(****************************************************************************************************<br>
© Syntegon Group.<br>
All rights reserved, also regarding any disposal, exploitation, reproduction, editing, distribution,<br>
as well as in the event of applications for industrial property rights.<br>
*****************************************************************************************************<br>
DESCRIPTION:<br>
Sets pose, track, strokes, gripper offsets and mover size. TRUE if anything changed.<br>
****************************************************************************************************)
METHOD m_Configure : BOOL
VAR_INPUT
	vi_Pose								: ST_VisuPose;	// MCS, track start on top of the movers with Z = 0
	vi_un_ModuleCount					: UINT;	// [-] track modules in a row
	vi_lr_ModuleLength					: LREAL;	// [mm]
	vi_lr_XMin							: LREAL;	// [mm]
	vi_lr_XMax							: LREAL;	// [mm]
	vi_lr_ZMin							: LREAL;	// [mm]
	vi_lr_ZMax							: LREAL;	// [mm]
	vi_lr_ToolOffsetX					: LREAL;	// [mm] gripper flange ahead of the X axis zero
	vi_lr_ToolOffsetZ					: LREAL;	// [mm] gripper flange relative to the mover top (below: negative)
	vi_lr_MoverLength					: LREAL;	// [mm] along the track
	vi_lr_MoverWidth					: LREAL;	// [mm]
END_VAR
VAR
	TempNew								: ST_VisuXtsGantryConfig;
END_VAR
TempNew := vo_Visu.stConfig;
TempNew.stPose := vi_Pose;
TempNew.nModuleCount := vi_un_ModuleCount;
TempNew.fModuleLength := vi_lr_ModuleLength;
TempNew.fXMin := vi_lr_XMin;
TempNew.fXMax := vi_lr_XMax;
TempNew.fZMin := vi_lr_ZMin;
TempNew.fZMax := vi_lr_ZMax;
TempNew.fToolOffsetX := vi_lr_ToolOffsetX;
TempNew.fToolOffsetZ := vi_lr_ToolOffsetZ;
TempNew.fMoverLength := vi_lr_MoverLength;
TempNew.fMoverWidth := vi_lr_MoverWidth;
m_Configure := m_ApplyConfig(TempNew);
END_METHOD

(****************************************************************************************************<br>
© Syntegon Group.<br>
All rights reserved, also regarding any disposal, exploitation, reproduction, editing, distribution,<br>
as well as in the event of applications for industrial property rights.<br>
*****************************************************************************************************<br>
DESCRIPTION:<br>
Sets or clears the fault of the whole gantry: drawn red with the message while active. Faults of single<br>
movers go through m_SetMover. The fault stays until it is cleared with m_SetFault(vi_b_Active := FALSE,<br>
vi_str_Message := ''). TRUE.<br>
****************************************************************************************************)
METHOD m_SetFault : BOOL
VAR_INPUT
	vi_b_Active							: BOOL;	// TRUE: fault active
	vi_str_Message						: STRING(80);	// shown to the operator; empty shows 'Fault'
END_VAR
vo_Visu.stState.stFault.bActive := vi_b_Active;
vo_Visu.stState.stFault.sMessage := vi_str_Message;
m_SetFault := TRUE;
END_METHOD

(****************************************************************************************************<br>
© Syntegon Group.<br>
All rights reserved, also regarding any disposal, exploitation, reproduction, editing, distribution,<br>
as well as in the event of applications for industrial property rights.<br>
*****************************************************************************************************<br>
DESCRIPTION:<br>
Defines finger vi_un_Finger (1-based) of every mover's gripper: a cylinder hanging from the finger's pose along<br>
its local -Z. The finger count grows to vi_un_Finger.<br>
*****************************************************************************************************<br>
OUTPUT VALUES:<br>
FALSE outside 1..VISU_GlobalConst_Param.VISU_un_MAX_FINGERS.<br>
****************************************************************************************************)
METHOD m_SetFinger : BOOL
VAR_INPUT
	vi_un_Finger						: UINT;	// [-] 1-based, as a product's nFingerId
	vi_lr_Diameter						: LREAL;	// [mm]
	vi_lr_Height						: LREAL;	// [mm] along the finger's local -Z
END_VAR
VAR
	TempNew								: ST_VisuXtsGantryConfig;
END_VAR
m_SetFinger := FALSE;
IF vi_un_Finger = 0 OR vi_un_Finger > VISU_GlobalConst_Param.VISU_un_MAX_FINGERS THEN
	RETURN;
END_IF
TempNew := vo_Visu.stConfig;
TempNew.aFingers[vi_un_Finger - 1].fDiameter := vi_lr_Diameter;
TempNew.aFingers[vi_un_Finger - 1].fHeight := vi_lr_Height;
TempNew.nFingerCount := MAX(TempNew.nFingerCount, vi_un_Finger);
m_ApplyConfig(TempNew);
m_SetFinger := TRUE;
END_METHOD

(****************************************************************************************************<br>
© Syntegon Group.<br>
All rights reserved, also regarding any disposal, exploitation, reproduction, editing, distribution,<br>
as well as in the event of applications for industrial property rights.<br>
*****************************************************************************************************<br>
DESCRIPTION:<br>
Reports one mover (actual values) at entry vi_un_Index and marks it valid. Call once per cycle per mover.<br>
*****************************************************************************************************<br>
OUTPUT VALUES:<br>
FALSE if vi_un_Index is outside the mover count set by m_SetMoverCount.<br>
****************************************************************************************************)
METHOD m_SetMover : BOOL
VAR_INPUT
	vi_un_Index							: UINT;	// [-] 0..m_SetMoverCount - 1
	vi_udn_Id							: UDINT;	// [-] unique within the gantry, > 0
	vi_lr_Position						: LREAL;	// [mm] along the track
	vi_lr_X								: LREAL;	// [mm] X axis
	vi_b_GripperActive					: BOOL;	// used only when no fingers are configured
	(* Finger poses absolute in the MCS and grip states, index 0 = finger 1; entries beyond the finger count are ignored. *)
	vi_FingerStates						: ARRAY[0..VISU_GlobalConst_Param.VISU_un_MAX_FINGERS - 1] OF ST_VisuFingerState;
	vi_b_Fault							: BOOL := FALSE;	// TRUE: this mover is in a fault
	vi_str_FaultMessage					: STRING(80) := '';	// shown to the operator; empty shows 'Fault'
END_VAR
m_SetMover := vi_un_Index < vo_Visu.stState.nMoverCount;
IF m_SetMover THEN
	vo_Visu.stState.aMovers[vi_un_Index].nId := vi_udn_Id;
	vo_Visu.stState.aMovers[vi_un_Index].bValid := TRUE;
	vo_Visu.stState.aMovers[vi_un_Index].fPosition := vi_lr_Position;
	vo_Visu.stState.aMovers[vi_un_Index].fX := vi_lr_X;
	vo_Visu.stState.aMovers[vi_un_Index].bGripperActive := vi_b_GripperActive;
	vo_Visu.stState.aMovers[vi_un_Index].aFingerStates := vi_FingerStates;
	vo_Visu.stState.aMovers[vi_un_Index].stFault.bActive := vi_b_Fault;
	vo_Visu.stState.aMovers[vi_un_Index].stFault.sMessage := vi_str_FaultMessage;
	vo_Visu.stState.nTimestamp := m_DcTime();
END_IF
END_METHOD

(****************************************************************************************************<br>
© Syntegon Group.<br>
All rights reserved, also regarding any disposal, exploitation, reproduction, editing, distribution,<br>
as well as in the event of applications for industrial property rights.<br>
*****************************************************************************************************<br>
DESCRIPTION:<br>
Sets how many mover entries are evaluated (limited to VISU_GlobalConst_Param.VISU_un_MAX_MOVERS); entries<br>
beyond are invalidated. TRUE if vi_un_Count fitted.<br>
****************************************************************************************************)
METHOD m_SetMoverCount : BOOL
VAR_INPUT
	vi_un_Count							: UINT;	// [-] movers
END_VAR
VAR
	un_TempIndex						: UINT;
END_VAR
m_SetMoverCount := vi_un_Count <= VISU_GlobalConst_Param.VISU_un_MAX_MOVERS;
vo_Visu.stState.nMoverCount := MIN(vi_un_Count, VISU_GlobalConst_Param.VISU_un_MAX_MOVERS);
FOR un_TempIndex := vo_Visu.stState.nMoverCount TO VISU_GlobalConst_Param.VISU_un_MAX_MOVERS - 1 DO
	vo_Visu.stState.aMovers[un_TempIndex].bValid := FALSE;
END_FOR
END_METHOD

(****************************************************************************************************<br>
© Syntegon Group.<br>
All rights reserved, also regarding any disposal, exploitation, reproduction, editing, distribution,<br>
as well as in the event of applications for industrial property rights.<br>
*****************************************************************************************************<br>
DESCRIPTION:<br>
Moves the gantry's shown coordinate system (origin triad, local measuring coordinates) away from the track<br>
start (stPose), in the gantry's local frame. Geometry and mover positions stay relative to stPose.<br>
TRUE if anything changed.<br>
****************************************************************************************************)
METHOD m_SetOriginShift : BOOL
VAR_INPUT
	vi_lr_X								: LREAL;	// [mm] along the gantry's local X
	vi_lr_Y								: LREAL := 0;	// [mm] along the track (local Y)
	vi_lr_Z								: LREAL := 0;	// [mm] along the gantry's local Z
END_VAR
VAR
	TempNew								: ST_VisuXtsGantryConfig;
END_VAR
TempNew := vo_Visu.stConfig;
TempNew.stOriginShift.fX := vi_lr_X;
TempNew.stOriginShift.fY := vi_lr_Y;
TempNew.stOriginShift.fZ := vi_lr_Z;
m_SetOriginShift := m_ApplyConfig(TempNew);
END_METHOD

(****************************************************************************************************<br>
© Syntegon Group.<br>
All rights reserved, also regarding any disposal, exploitation, reproduction, editing, distribution,<br>
as well as in the event of applications for industrial property rights.<br>
*****************************************************************************************************<br>
DESCRIPTION:<br>
Adds a pick or place zone, or updates the one for the same conveyor and kind.<br>
*****************************************************************************************************<br>
OUTPUT VALUES:<br>
FALSE for vi_udn_ConveyorId = 0 or a full list.<br>
****************************************************************************************************)
METHOD m_SetZone : BOOL
VAR_INPUT
	vi_udn_ConveyorId					: UDINT;	// [-] manifest id of the conveyor
	vi_e_Kind							: E_VisuZoneKind;
	vi_lr_Start							: LREAL;	// [mm] along the conveyor from its origin (belt coordinates, not MCS)
	vi_lr_End							: LREAL;	// [mm] along the conveyor from its origin
	vi_lr_AllocationOffset				: LREAL := 0;	// [mm] before vi_lr_End up to which products may be allocated; 0 = no limit
	vi_lr_CcsOffset						: LREAL := 0;	// [mm] along the conveyor from its origin: the robot's conveyor coordinate system
END_VAR
VAR
	TempNew								: ST_VisuXtsGantryConfig;
	un_TempIndex						: UINT;
END_VAR
m_SetZone := FALSE;
IF vi_udn_ConveyorId = 0 THEN
	RETURN;
END_IF
TempNew := vo_Visu.stConfig;
un_TempIndex := 0;
(* ST evaluates both operands of AND: test the index before reading the array. *)
WHILE un_TempIndex < TempNew.nZoneCount DO
	IF TempNew.aZones[un_TempIndex].nConveyorId = vi_udn_ConveyorId AND TempNew.aZones[un_TempIndex].eKind = vi_e_Kind THEN
		EXIT;
	END_IF
	un_TempIndex := un_TempIndex + 1;
END_WHILE
IF un_TempIndex >= VISU_GlobalConst_Param.VISU_un_MAX_ZONES THEN
	RETURN;
END_IF
IF un_TempIndex = TempNew.nZoneCount THEN
	TempNew.nZoneCount := TempNew.nZoneCount + 1;
END_IF
TempNew.aZones[un_TempIndex].nConveyorId := vi_udn_ConveyorId;
TempNew.aZones[un_TempIndex].eKind := vi_e_Kind;
TempNew.aZones[un_TempIndex].fStart := vi_lr_Start;
TempNew.aZones[un_TempIndex].fEnd := vi_lr_End;
TempNew.aZones[un_TempIndex].fAllocationOffset := vi_lr_AllocationOffset;
TempNew.aZones[un_TempIndex].fCcsOffset := vi_lr_CcsOffset;
m_ApplyConfig(TempNew);
m_SetZone := TRUE;
END_METHOD

(****************************************************************************************************<br>
© Syntegon Group.<br>
All rights reserved, also regarding any disposal, exploitation, reproduction, editing, distribution,<br>
as well as in the event of applications for industrial property rights.<br>
*****************************************************************************************************<br>
DESCRIPTION:<br>
Reports the common Z axis (actual value). Call once per cycle; it also stamps the state with the cycle's DC time.<br>
****************************************************************************************************)
METHOD m_SetZPosition : BOOL
VAR_INPUT
	vi_lr_Z								: LREAL;	// [mm]
END_VAR
vo_Visu.stState.fZ := vi_lr_Z;
vo_Visu.stState.nTimestamp := m_DcTime();
m_SetZPosition := TRUE;
END_METHOD

END_FUNCTION_BLOCK

// POUs/_FB_VisuXtsLoop
(****************************************************************************************************<br>
© Syntegon Group.<br>
All rights reserved, also regarding any disposal, exploitation, reproduction, editing, distribution,<br>
as well as in the event of applications for industrial property rights.<br>
*****************************************************************************************************<br>
DESCRIPTION:<br>
One visualised XTS loop (e.g. Fxx): movers circulating on a closed track of two straights and two 180 deg curves.<br>
Typical cycle:<br>
  fb_Fxx.m_Register(vio_Manifest := GVL_Visu.stManifest, vi_udn_Id := 20, vi_str_Name := 'Fxx',<br>
      vi_str_Path := 'MAIN.fb_Fxx.vo_Visu');<br>
  fb_Fxx.m_Configure(vi_Pose := LoopPose, vi_lr_StraightLength := 2400, vi_lr_CurveRadius := 250,<br>
      vi_lr_ToolOffset := 120, vi_lr_MoverLength := 100, vi_lr_MoverWidth := 60);<br>
  fb_Fxx.m_SetFinger(vi_un_Finger := 1, vi_lr_Diameter := 40, vi_lr_Height := 50);<br>
  fb_Fxx.m_SetZone(vi_udn_ConveyorId := 2, vi_e_Kind := E_VisuZoneKind.PICK, vi_lr_Start := 2200, vi_lr_End := 2800);<br>
  fb_Fxx.m_SetMoverCount(12);<br>
  fb_Fxx.m_SetMover(vi_un_Index := 0, vi_udn_Id := 1, vi_lr_Position := ..., vi_FingerStates := Mover1Fingers);<br>
Positions run along the loop from the start of the lower straight in the conveying direction (0..m_Perimeter()).<br>
The config methods may be called every cycle; the config version only changes when a value does.<br>
*****************************************************************************************************<br>
OUTPUT VALUES:<br>
vo_Visu is the contract structure the gateway reads at the path given to m_Register. Do not write it.<br>
*****************************************************************************************************<br>
VERSION         ¦ DATE       ¦ NAME      ¦ CHANGE<br>
Syn_Visu 3.0.0  ¦ 2026-10-31 ¦ J.Willner ¦ Naming and layout after the TCAT programming guideline<br>
****************************************************************************************************)
FUNCTION_BLOCK _FB_VisuXtsLoop EXTENDS _FB_VisuComponent
VAR_OUTPUT
	vo_Visu								: ST_VisuXtsLoop;	// contract structure read by the gateway
END_VAR

(****************************************************************************************************<br>
© Syntegon Group.<br>
All rights reserved, also regarding any disposal, exploitation, reproduction, editing, distribution,<br>
as well as in the event of applications for industrial property rights.<br>
*****************************************************************************************************<br>
DESCRIPTION:<br>
Takes over vio_New and increments the config version if it differs from the current config. TRUE if changed.<br>
****************************************************************************************************)
METHOD PRIVATE m_ApplyConfig : BOOL
VAR_IN_OUT
	vio_New								: ST_VisuXtsLoopConfig;
END_VAR
m_ApplyConfig := Tc2_System.MEMCMP(ADR(vio_New), ADR(vo_Visu.stConfig), SIZEOF(vio_New)) <> 0;
IF m_ApplyConfig THEN
	vo_Visu.stConfig := vio_New;
	m_NotifyConfigChanged();
END_IF
END_METHOD

(****************************************************************************************************<br>
© Syntegon Group.<br>
All rights reserved, also regarding any disposal, exploitation, reproduction, editing, distribution,<br>
as well as in the event of applications for industrial property rights.<br>
*****************************************************************************************************<br>
DESCRIPTION:<br>
Removes the gripper definition. TRUE if there was one.<br>
****************************************************************************************************)
METHOD m_ClearFingers : BOOL
VAR
	TempNew								: ST_VisuXtsLoopConfig;
	TempEmpty							: ST_VisuFinger;
	un_TempIndex						: UINT;
END_VAR
TempNew := vo_Visu.stConfig;
FOR un_TempIndex := 0 TO VISU_GlobalConst_Param.VISU_un_MAX_FINGERS - 1 DO
	TempNew.aFingers[un_TempIndex] := TempEmpty;
END_FOR
TempNew.nFingerCount := 0;
m_ClearFingers := m_ApplyConfig(TempNew);
END_METHOD

(****************************************************************************************************<br>
© Syntegon Group.<br>
All rights reserved, also regarding any disposal, exploitation, reproduction, editing, distribution,<br>
as well as in the event of applications for industrial property rights.<br>
*****************************************************************************************************<br>
DESCRIPTION:<br>
Removes all pick and place zones. TRUE if there were any.<br>
****************************************************************************************************)
METHOD m_ClearZones : BOOL
VAR
	TempNew								: ST_VisuXtsLoopConfig;
	TempEmpty							: ST_VisuZone;
	un_TempIndex						: UINT;
END_VAR
TempNew := vo_Visu.stConfig;
FOR un_TempIndex := 0 TO VISU_GlobalConst_Param.VISU_un_MAX_ZONES - 1 DO
	TempNew.aZones[un_TempIndex] := TempEmpty;
END_FOR
TempNew.nZoneCount := 0;
m_ClearZones := m_ApplyConfig(TempNew);
END_METHOD

(****************************************************************************************************<br>
© Syntegon Group.<br>
All rights reserved, also regarding any disposal, exploitation, reproduction, editing, distribution,<br>
as well as in the event of applications for industrial property rights.<br>
*****************************************************************************************************<br>
DESCRIPTION:<br>
Manifest type: XTS loop.<br>
****************************************************************************************************)
METHOD PROTECTED m_ComponentType : E_VisuComponentType
m_ComponentType := E_VisuComponentType.XTS_LOOP;
END_METHOD

(****************************************************************************************************<br>
© Syntegon Group.<br>
All rights reserved, also regarding any disposal, exploitation, reproduction, editing, distribution,<br>
as well as in the event of applications for industrial property rights.<br>
*****************************************************************************************************<br>
DESCRIPTION:<br>
Sets pose, track geometry, tool offset and mover size. TRUE if anything changed.<br>
****************************************************************************************************)
METHOD m_Configure : BOOL
VAR_INPUT
	vi_Pose								: ST_VisuPose;	// MCS, start of the lower straight; the loop stands in the local X-Z plane
	vi_lr_StraightLength				: LREAL;	// [mm]
	vi_lr_CurveRadius					: LREAL;	// [mm]
	vi_lr_ToolOffset					: LREAL;	// [mm] tool point outwards from the track
	vi_lr_MoverLength					: LREAL;	// [mm] along the track
	vi_lr_MoverWidth					: LREAL;	// [mm]
END_VAR
VAR
	TempNew								: ST_VisuXtsLoopConfig;
END_VAR
TempNew := vo_Visu.stConfig;
TempNew.stPose := vi_Pose;
TempNew.fStraightLength := vi_lr_StraightLength;
TempNew.fCurveRadius := vi_lr_CurveRadius;
TempNew.fToolOffset := vi_lr_ToolOffset;
TempNew.fMoverLength := vi_lr_MoverLength;
TempNew.fMoverWidth := vi_lr_MoverWidth;
m_Configure := m_ApplyConfig(TempNew);
END_METHOD

(****************************************************************************************************<br>
© Syntegon Group.<br>
All rights reserved, also regarding any disposal, exploitation, reproduction, editing, distribution,<br>
as well as in the event of applications for industrial property rights.<br>
*****************************************************************************************************<br>
DESCRIPTION:<br>
Length of the loop as the visualisation computes it (curves as semicircles), [mm].<br>
****************************************************************************************************)
METHOD m_Perimeter : LREAL
m_Perimeter := 2.0 * vo_Visu.stConfig.fStraightLength + 2.0 * 3.141592653589793 * vo_Visu.stConfig.fCurveRadius;
END_METHOD

(****************************************************************************************************<br>
© Syntegon Group.<br>
All rights reserved, also regarding any disposal, exploitation, reproduction, editing, distribution,<br>
as well as in the event of applications for industrial property rights.<br>
*****************************************************************************************************<br>
DESCRIPTION:<br>
Sets or clears the fault of the whole loop: drawn red with the message while active. Faults of single<br>
movers go through m_SetMover. The fault stays until it is cleared with m_SetFault(vi_b_Active := FALSE,<br>
vi_str_Message := ''). TRUE.<br>
****************************************************************************************************)
METHOD m_SetFault : BOOL
VAR_INPUT
	vi_b_Active							: BOOL;	// TRUE: fault active
	vi_str_Message						: STRING(80);	// shown to the operator; empty shows 'Fault'
END_VAR
vo_Visu.stState.stFault.bActive := vi_b_Active;
vo_Visu.stState.stFault.sMessage := vi_str_Message;
m_SetFault := TRUE;
END_METHOD

(****************************************************************************************************<br>
© Syntegon Group.<br>
All rights reserved, also regarding any disposal, exploitation, reproduction, editing, distribution,<br>
as well as in the event of applications for industrial property rights.<br>
*****************************************************************************************************<br>
DESCRIPTION:<br>
Defines finger vi_un_Finger (1-based) of every mover's gripper: a cylinder hanging from the finger's pose along<br>
its local -Z. The finger count grows to vi_un_Finger.<br>
*****************************************************************************************************<br>
OUTPUT VALUES:<br>
FALSE outside 1..VISU_GlobalConst_Param.VISU_un_MAX_FINGERS.<br>
****************************************************************************************************)
METHOD m_SetFinger : BOOL
VAR_INPUT
	vi_un_Finger						: UINT;	// [-] 1-based, as a product's nFingerId
	vi_lr_Diameter						: LREAL;	// [mm]
	vi_lr_Height						: LREAL;	// [mm] along the finger's local -Z
END_VAR
VAR
	TempNew								: ST_VisuXtsLoopConfig;
END_VAR
m_SetFinger := FALSE;
IF vi_un_Finger = 0 OR vi_un_Finger > VISU_GlobalConst_Param.VISU_un_MAX_FINGERS THEN
	RETURN;
END_IF
TempNew := vo_Visu.stConfig;
TempNew.aFingers[vi_un_Finger - 1].fDiameter := vi_lr_Diameter;
TempNew.aFingers[vi_un_Finger - 1].fHeight := vi_lr_Height;
TempNew.nFingerCount := MAX(TempNew.nFingerCount, vi_un_Finger);
m_ApplyConfig(TempNew);
m_SetFinger := TRUE;
END_METHOD

(****************************************************************************************************<br>
© Syntegon Group.<br>
All rights reserved, also regarding any disposal, exploitation, reproduction, editing, distribution,<br>
as well as in the event of applications for industrial property rights.<br>
*****************************************************************************************************<br>
DESCRIPTION:<br>
Reports one mover at entry vi_un_Index and marks it valid. Call once per cycle per mover.<br>
*****************************************************************************************************<br>
OUTPUT VALUES:<br>
FALSE if vi_un_Index is outside the mover count set by m_SetMoverCount.<br>
****************************************************************************************************)
METHOD m_SetMover : BOOL
VAR_INPUT
	vi_un_Index							: UINT;	// [-] 0..m_SetMoverCount - 1
	vi_udn_Id							: UDINT;	// [-] unique within the loop, > 0
	vi_lr_Position						: LREAL;	// [mm] along the loop from the start of the lower straight (0..m_Perimeter())
	(* Finger poses absolute in the MCS and grip states, index 0 = finger 1; entries beyond the finger count are ignored. *)
	vi_FingerStates						: ARRAY[0..VISU_GlobalConst_Param.VISU_un_MAX_FINGERS - 1] OF ST_VisuFingerState;
	vi_b_Fault							: BOOL := FALSE;	// TRUE: this mover is in a fault
	vi_str_FaultMessage					: STRING(80) := '';	// shown to the operator; empty shows 'Fault'
END_VAR
m_SetMover := vi_un_Index < vo_Visu.stState.nMoverCount;
IF m_SetMover THEN
	vo_Visu.stState.aMovers[vi_un_Index].nId := vi_udn_Id;
	vo_Visu.stState.aMovers[vi_un_Index].bValid := TRUE;
	vo_Visu.stState.aMovers[vi_un_Index].fPosition := vi_lr_Position;
	vo_Visu.stState.aMovers[vi_un_Index].aFingerStates := vi_FingerStates;
	vo_Visu.stState.aMovers[vi_un_Index].stFault.bActive := vi_b_Fault;
	vo_Visu.stState.aMovers[vi_un_Index].stFault.sMessage := vi_str_FaultMessage;
	vo_Visu.stState.nTimestamp := m_DcTime();
END_IF
END_METHOD

(****************************************************************************************************<br>
© Syntegon Group.<br>
All rights reserved, also regarding any disposal, exploitation, reproduction, editing, distribution,<br>
as well as in the event of applications for industrial property rights.<br>
*****************************************************************************************************<br>
DESCRIPTION:<br>
Sets how many mover entries are evaluated (limited to VISU_GlobalConst_Param.VISU_un_MAX_MOVERS); entries<br>
beyond are invalidated. TRUE if vi_un_Count fitted.<br>
****************************************************************************************************)
METHOD m_SetMoverCount : BOOL
VAR_INPUT
	vi_un_Count							: UINT;	// [-] movers
END_VAR
VAR
	un_TempIndex						: UINT;
END_VAR
m_SetMoverCount := vi_un_Count <= VISU_GlobalConst_Param.VISU_un_MAX_MOVERS;
vo_Visu.stState.nMoverCount := MIN(vi_un_Count, VISU_GlobalConst_Param.VISU_un_MAX_MOVERS);
FOR un_TempIndex := vo_Visu.stState.nMoverCount TO VISU_GlobalConst_Param.VISU_un_MAX_MOVERS - 1 DO
	vo_Visu.stState.aMovers[un_TempIndex].bValid := FALSE;
END_FOR
END_METHOD

(****************************************************************************************************<br>
© Syntegon Group.<br>
All rights reserved, also regarding any disposal, exploitation, reproduction, editing, distribution,<br>
as well as in the event of applications for industrial property rights.<br>
*****************************************************************************************************<br>
DESCRIPTION:<br>
Moves the loop's shown coordinate system (origin triad, local measuring coordinates) away from the start of<br>
the lower straight (stPose), in the loop's local frame. Geometry and mover positions stay relative to stPose.<br>
TRUE if anything changed.<br>
****************************************************************************************************)
METHOD m_SetOriginShift : BOOL
VAR_INPUT
	vi_lr_X								: LREAL;	// [mm] along the lower straight (local X)
	vi_lr_Y								: LREAL := 0;	// [mm] along the loop's local Y
	vi_lr_Z								: LREAL := 0;	// [mm] along the loop's local Z
END_VAR
VAR
	TempNew								: ST_VisuXtsLoopConfig;
END_VAR
TempNew := vo_Visu.stConfig;
TempNew.stOriginShift.fX := vi_lr_X;
TempNew.stOriginShift.fY := vi_lr_Y;
TempNew.stOriginShift.fZ := vi_lr_Z;
m_SetOriginShift := m_ApplyConfig(TempNew);
END_METHOD

(****************************************************************************************************<br>
© Syntegon Group.<br>
All rights reserved, also regarding any disposal, exploitation, reproduction, editing, distribution,<br>
as well as in the event of applications for industrial property rights.<br>
*****************************************************************************************************<br>
DESCRIPTION:<br>
Adds a pick or place zone, or updates the one for the same conveyor and kind.<br>
*****************************************************************************************************<br>
OUTPUT VALUES:<br>
FALSE for vi_udn_ConveyorId = 0 or a full list.<br>
****************************************************************************************************)
METHOD m_SetZone : BOOL
VAR_INPUT
	vi_udn_ConveyorId					: UDINT;	// [-] manifest id of the conveyor
	vi_e_Kind							: E_VisuZoneKind;
	vi_lr_Start							: LREAL;	// [mm] along the conveyor from its origin (belt coordinates, not MCS)
	vi_lr_End							: LREAL;	// [mm] along the conveyor from its origin
	vi_lr_AllocationOffset				: LREAL := 0;	// [mm] before vi_lr_End up to which products may be allocated; 0 = no limit
	vi_lr_CcsOffset						: LREAL := 0;	// [mm] along the conveyor from its origin: the robot's conveyor coordinate system
END_VAR
VAR
	TempNew								: ST_VisuXtsLoopConfig;
	un_TempIndex						: UINT;
END_VAR
m_SetZone := FALSE;
IF vi_udn_ConveyorId = 0 THEN
	RETURN;
END_IF
TempNew := vo_Visu.stConfig;
un_TempIndex := 0;
(* ST evaluates both operands of AND: test the index before reading the array. *)
WHILE un_TempIndex < TempNew.nZoneCount DO
	IF TempNew.aZones[un_TempIndex].nConveyorId = vi_udn_ConveyorId AND TempNew.aZones[un_TempIndex].eKind = vi_e_Kind THEN
		EXIT;
	END_IF
	un_TempIndex := un_TempIndex + 1;
END_WHILE
IF un_TempIndex >= VISU_GlobalConst_Param.VISU_un_MAX_ZONES THEN
	RETURN;
END_IF
IF un_TempIndex = TempNew.nZoneCount THEN
	TempNew.nZoneCount := TempNew.nZoneCount + 1;
END_IF
TempNew.aZones[un_TempIndex].nConveyorId := vi_udn_ConveyorId;
TempNew.aZones[un_TempIndex].eKind := vi_e_Kind;
TempNew.aZones[un_TempIndex].fStart := vi_lr_Start;
TempNew.aZones[un_TempIndex].fEnd := vi_lr_End;
TempNew.aZones[un_TempIndex].fAllocationOffset := vi_lr_AllocationOffset;
TempNew.aZones[un_TempIndex].fCcsOffset := vi_lr_CcsOffset;
m_ApplyConfig(TempNew);
m_SetZone := TRUE;
END_METHOD

END_FUNCTION_BLOCK

// POUs/_FC_GetVersionSynVisu
(****************************************************************************************************<br>
© Syntegon Group.<br>
All rights reserved, also regarding any disposal, exploitation, reproduction, editing, distribution,<br>
as well as in the event of applications for industrial property rights.<br>
*****************************************************************************************************<br>
DESCRIPTION:<br>
Runtime-readable version of the Syn_Visu library.<br>
*****************************************************************************************************<br>
VERSION         ¦ DATE       ¦ NAME      ¦ CHANGE<br>
Syn_Visu 3.0.0  ¦ 2026-10-31 ¦ J.Willner ¦ Naming and layout after the TCAT programming guideline<br>
Syn_Visu 3.1.0  ¦ 2026-10-31 ¦ J.Willner ¦ Faults of components and XTS movers (protocol 8)<br>
Syn_Visu 3.2.0  ¦ 2026-10-31 ¦ J.Willner ¦ _FB_VisuConveyor.m_MoveProduct<br>
Syn_Visu 3.3.0  ¦ 2026-10-31 ¦ J.Willner ¦ Zone CCS offset, origin shift per component (protocol 9)<br>
****************************************************************************************************)
FUNCTION _FC_GetVersionSynVisu : UINT
VAR_INPUT
	vi_n_VersionElement					: INT;	// [-] 1 = major, 2 = minor, 3 = revision
END_VAR

CASE vi_n_VersionElement OF
	1: _FC_GetVersionSynVisu := 3;
	2: _FC_GetVersionSynVisu := 3;
	3: _FC_GetVersionSynVisu := 0;
ELSE
	_FC_GetVersionSynVisu := 16#FFFF;
END_CASE

END_FUNCTION
